// SIMATIC S7-200 SMART project (STEP 7-Micro/WIN SMART), CPU ST40

SYMBOL_TABLE System Symbols
ON_STATE         M0.0     // ON STATE
END_SYMBOL_TABLE

SYMBOL_TABLE STEPS MEMORY
PROCESS          M1.0     // PROCESS
STEP_1_DONE      M1.1     // STEP_1_DONE
STEP_2_DONE      M1.2     // STEP_2_DONE
STEP_3_DONE      M1.3     // STEP_3_DONE
STEP_4_DONE      M1.4     // STEP_4_DONE
STEP_5_DONE      M1.5     // STEP_5_DONE
STEP_6_DONE      M1.6     // STEP_6_DONE
STEP_7_DONE      M1.7     // STEP_7_DONE
STEP_8_DONE      M2.0     // STEP_8_DONE
STEP_9_DONE      M2.1     // STEP_9_DONE
STEP_10_DONE     M2.2     // STEP_10_DONE
STEP_11_DONE     M2.3     // STEP_11_DONE
STEP_12_DONE     M2.4     // STEP_12_DONE
END_SYMBOL_TABLE

SYMBOL_TABLE MOVEMENT MEMORY
X_MOVEMENT       M3.0     // X_MOVEMENT
Y_MOVEMENT       M3.1     // Y_MOVEMENT
Z_MOVEMENT       M3.2     // Z_MOVEMENT
GRIPPER_MOVEMENT M3.3     // GRIPPER_MOVEMENT
END_SYMBOL_TABLE

ORGANIZATION_BLOCK MAIN:OB1
TITLE=Program Comments
BEGIN
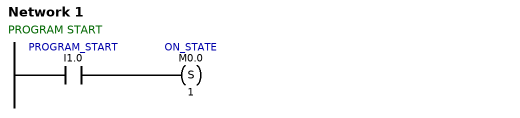
Network 1
// PROGRAM START
LD     PROGRAM_START:I1.0
S      ON_STATE:M0.0, 1
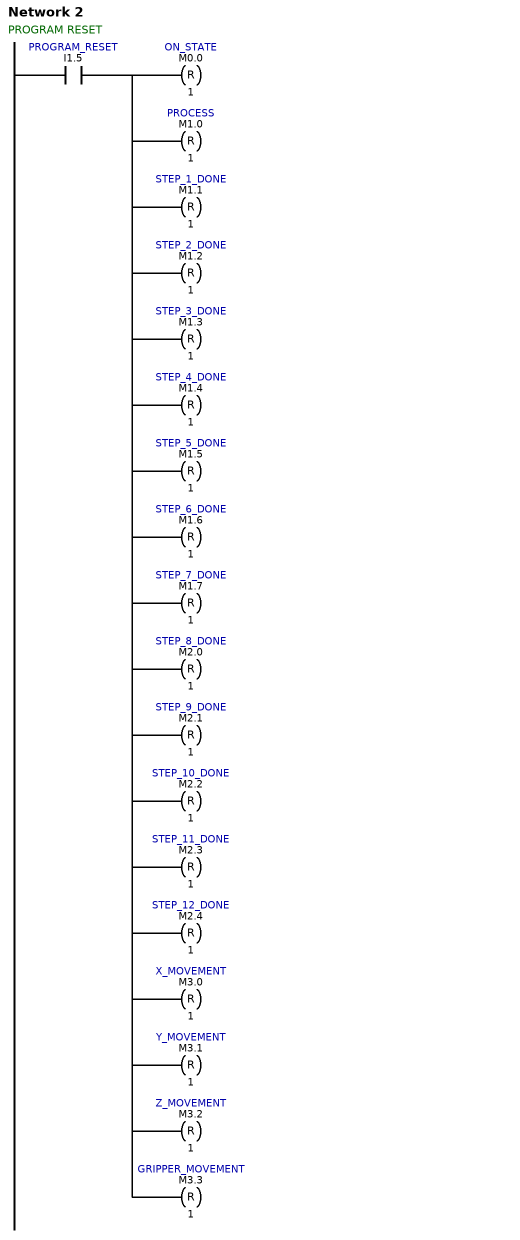
Network 2
// PROGRAM RESET
LD     PROGRAM_RESET:I1.5
R      ON_STATE:M0.0, 1
R      PROCESS:M1.0, 1
R      STEP_1_DONE:M1.1, 1
R      STEP_2_DONE:M1.2, 1
R      STEP_3_DONE:M1.3, 1
R      STEP_4_DONE:M1.4, 1
R      STEP_5_DONE:M1.5, 1
R      STEP_6_DONE:M1.6, 1
R      STEP_7_DONE:M1.7, 1
R      STEP_8_DONE:M2.0, 1
R      STEP_9_DONE:M2.1, 1
R      STEP_10_DONE:M2.2, 1
R      STEP_11_DONE:M2.3, 1
R      STEP_12_DONE:M2.4, 1
R      X_MOVEMENT:M3.0, 1
R      Y_MOVEMENT:M3.1, 1
R      Z_MOVEMENT:M3.2, 1
R      GRIPPER_MOVEMENT:M3.3, 1
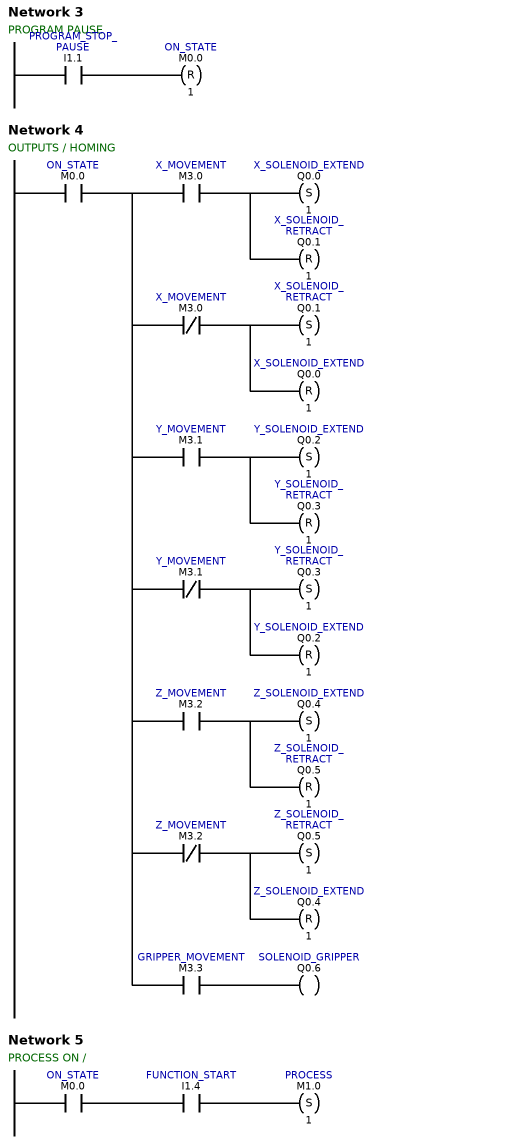
Network 3
// PROGRAM PAUSE
LD     PROGRAM_STOP_PAUSE:I1.1
R      ON_STATE:M0.0, 1
Network 4
// OUTPUTS / HOMING
LD     ON_STATE:M0.0
LPS
A      X_MOVEMENT:M3.0
S      X_SOLENOID_EXTEND:Q0.0, 1
R      X_SOLENOID_RETRACT:Q0.1, 1
LRD
AN     X_MOVEMENT:M3.0
S      X_SOLENOID_RETRACT:Q0.1, 1
R      X_SOLENOID_EXTEND:Q0.0, 1
LRD
A      Y_MOVEMENT:M3.1
S      Y_SOLENOID_EXTEND:Q0.2, 1
R      Y_SOLENOID_RETRACT:Q0.3, 1
LRD
AN     Y_MOVEMENT:M3.1
S      Y_SOLENOID_RETRACT:Q0.3, 1
R      Y_SOLENOID_EXTEND:Q0.2, 1
LRD
A      Z_MOVEMENT:M3.2
S      Z_SOLENOID_EXTEND:Q0.4, 1
R      Z_SOLENOID_RETRACT:Q0.5, 1
LRD
AN     Z_MOVEMENT:M3.2
S      Z_SOLENOID_RETRACT:Q0.5, 1
R      Z_SOLENOID_EXTEND:Q0.4, 1
LPP
A      GRIPPER_MOVEMENT:M3.3
=      SOLENOID_GRIPPER:Q0.6
Network 5
// PROCESS ON
// 
LD     ON_STATE:M0.0
A      FUNCTION_START:I1.4
S      PROCESS:M1.0, 1
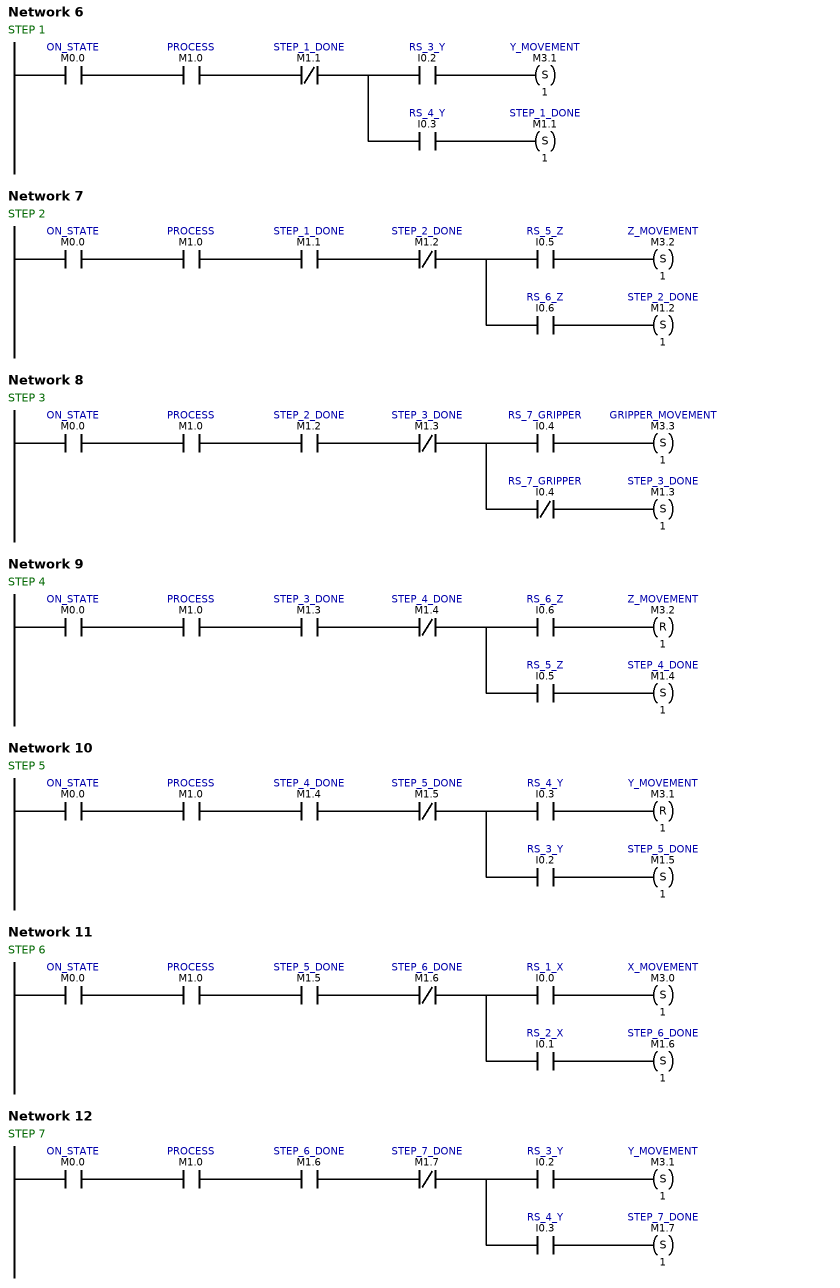
Network 6
// STEP 1 
LD     ON_STATE:M0.0
A      PROCESS:M1.0
AN     STEP_1_DONE:M1.1
LPS
A      RS_3_Y:I0.2
S      Y_MOVEMENT:M3.1, 1
LPP
A      RS_4_Y:I0.3
S      STEP_1_DONE:M1.1, 1
Network 7
// STEP 2 
LD     ON_STATE:M0.0
A      PROCESS:M1.0
A      STEP_1_DONE:M1.1
AN     STEP_2_DONE:M1.2
LPS
A      RS_5_Z:I0.5
S      Z_MOVEMENT:M3.2, 1
LPP
A      RS_6_Z:I0.6
S      STEP_2_DONE:M1.2, 1
Network 8
// STEP 3 
LD     ON_STATE:M0.0
A      PROCESS:M1.0
A      STEP_2_DONE:M1.2
AN     STEP_3_DONE:M1.3
LPS
A      RS_7_GRIPPER:I0.4
S      GRIPPER_MOVEMENT:M3.3, 1
LPP
AN     RS_7_GRIPPER:I0.4
S      STEP_3_DONE:M1.3, 1
Network 9
// STEP 4
LD     ON_STATE:M0.0
A      PROCESS:M1.0
A      STEP_3_DONE:M1.3
AN     STEP_4_DONE:M1.4
LPS
A      RS_6_Z:I0.6
R      Z_MOVEMENT:M3.2, 1
LPP
A      RS_5_Z:I0.5
S      STEP_4_DONE:M1.4, 1
Network 10
// STEP 5
LD     ON_STATE:M0.0
A      PROCESS:M1.0
A      STEP_4_DONE:M1.4
AN     STEP_5_DONE:M1.5
LPS
A      RS_4_Y:I0.3
R      Y_MOVEMENT:M3.1, 1
LPP
A      RS_3_Y:I0.2
S      STEP_5_DONE:M1.5, 1
Network 11
// STEP 6
LD     ON_STATE:M0.0
A      PROCESS:M1.0
A      STEP_5_DONE:M1.5
AN     STEP_6_DONE:M1.6
LPS
A      RS_1_X:I0.0
S      X_MOVEMENT:M3.0, 1
LPP
A      RS_2_X:I0.1
S      STEP_6_DONE:M1.6, 1
Network 12
// STEP 7
LD     ON_STATE:M0.0
A      PROCESS:M1.0
A      STEP_6_DONE:M1.6
AN     STEP_7_DONE:M1.7
LPS
A      RS_3_Y:I0.2
S      Y_MOVEMENT:M3.1, 1
LPP
A      RS_4_Y:I0.3
S      STEP_7_DONE:M1.7, 1
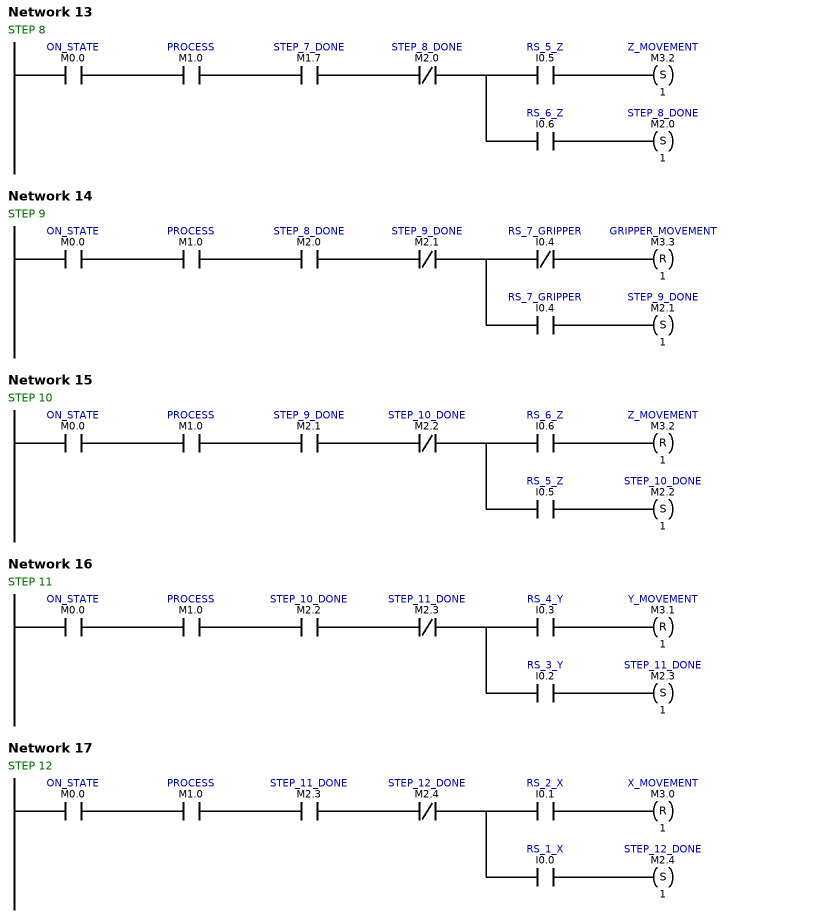
Network 13
// STEP 8
LD     ON_STATE:M0.0
A      PROCESS:M1.0
A      STEP_7_DONE:M1.7
AN     STEP_8_DONE:M2.0
LPS
A      RS_5_Z:I0.5
S      Z_MOVEMENT:M3.2, 1
LPP
A      RS_6_Z:I0.6
S      STEP_8_DONE:M2.0, 1
Network 14
// STEP 9
LD     ON_STATE:M0.0
A      PROCESS:M1.0
A      STEP_8_DONE:M2.0
AN     STEP_9_DONE:M2.1
LPS
AN     RS_7_GRIPPER:I0.4
R      GRIPPER_MOVEMENT:M3.3, 1
LPP
A      RS_7_GRIPPER:I0.4
S      STEP_9_DONE:M2.1, 1
Network 15
// STEP 10
LD     ON_STATE:M0.0
A      PROCESS:M1.0
A      STEP_9_DONE:M2.1
AN     STEP_10_DONE:M2.2
LPS
A      RS_6_Z:I0.6
R      Z_MOVEMENT:M3.2, 1
LPP
A      RS_5_Z:I0.5
S      STEP_10_DONE:M2.2, 1
Network 16
// STEP 11
LD     ON_STATE:M0.0
A      PROCESS:M1.0
A      STEP_10_DONE:M2.2
AN     STEP_11_DONE:M2.3
LPS
A      RS_4_Y:I0.3
R      Y_MOVEMENT:M3.1, 1
LPP
A      RS_3_Y:I0.2
S      STEP_11_DONE:M2.3, 1
Network 17
// STEP 12
LD     ON_STATE:M0.0
A      PROCESS:M1.0
A      STEP_11_DONE:M2.3
AN     STEP_12_DONE:M2.4
LPS
A      RS_2_X:I0.1
R      X_MOVEMENT:M3.0, 1
LPP
A      RS_1_X:I0.0
S      STEP_12_DONE:M2.4, 1
END_ORGANIZATION_BLOCK
